// TIA Portal V21 export
PlcForceTable "Force table"
  PlcForceTableEntry ""Valve":P"  DisplayFormat=Bool, MonitorTrigger=Permanent, Comment="Keep the inlet open"
  PlcForceTableEntry ""DoorClosed":P"  DisplayFormat=Bool, MonitorTrigger=Permanent
